FUNCTION_BLOCK FB_BOSCH_DriveLink
VAR_INPUT
	pDrive							:POINTER TO ST_BOSCHINDRADRIVECIA402_REF;			(* The DRIVE_REF data type  is an interface between the PLC and the DRIVE and contains axis information *)
END_VAR
VAR_OUTPUT		

END_VAR
VAR_IN_OUT

END_VAR
VAR
END_VAR


	
pDrive^.bDriverZKL3 := pDrive^.stBoschToPlc.wDriveStatuswordS00135.11;			(* Drive change bit class 3 diagnostics *)
pDrive^.bDriverZKL2 := pDrive^.stBoschToPlc.wDriveStatuswordS00135.12;			(* Drive change bit class 2 diagnostics *)
pDrive^.bDriverZKL1 := pDrive^.stBoschToPlc.wDriveStatuswordS00135.13;			(* Drive error, error in class 1 diagnostics *)
	
pDrive^.bDriveBB :=	pDrive^.stBoschToPlc.wDriveStatuswordS00135.14				(* Drive ready for power on *)
					AND NOT pDrive^.stBoschToPlc.wDriveStatuswordS00135.15;
pDrive^.bDriveAB :=	NOT pDrive^.stBoschToPlc.wDriveStatuswordS00135.14			(* Drive control section and power section ready for operation, torque-free*)
					AND pDrive^.stBoschToPlc.wDriveStatuswordS00135.15;
pDrive^.bDriveAF :=	pDrive^.stBoschToPlc.wDriveStatuswordS00135.14				(* Drive in operation, with torque *)
					AND pDrive^.stBoschToPlc.wDriveStatuswordS00135.15;

END_FUNCTION_BLOCK

(* stored: Version 1.1.0.1, ProductVersion 3.1.4024.15
   POU FB_BOSCH_DriveLink: Id {7b25cd81-1b2d-47fe-a7a5-f97947ab44ab}, SpecialFunc None *)
